Fanuc KAREL source: ka00142.KL

PROGRAM KA00142
%STACKSIZE=65535
%PRIORITY=65535
%NOLOCKGROUP
VAR
SRC : ARRAY[2] OF SHORT
-- UNRESOLVED DECLARATIONS (source type spelling not recovered)
-- DST : TYPE_0x001C (type_u16=0x001C)
BEGIN
SRC[1]=2
DST=SRC[1]
END KA00142
